// Lecture brute d'une entrée analogique (docs/04 § 6.1) : référence invalide -> 0
FUNCTION F_ReadAI : INT
VAR_INPUT
    stRef : ST_SignalRef;
END_VAR

IF stRef.eKind <> E_SignalKind.AI OR GVL_IoRef.pAI = 0 OR stRef.nIndex < 0 OR stRef.nIndex >= GVL_Const.MAX_AI THEN
    F_ReadAI := 0;
    RETURN;
END_IF
F_ReadAI := GVL_IoRef.pAI^[stRef.nIndex];

END_FUNCTION

(* stored: Version 1.1.0.1, ProductVersion 3.1.4024.12
   POU F_ReadAI: Id {92c952a7-9e34-5907-a605-4df56dabecd5}, SpecialFunc None *)
